// Mock of FB_AzimuthControl for the telescope state machine tests (MONETcommon#36, BROTLib plan 2026-10-21-telescope-state-machine-unification D1).
FUNCTION_BLOCK FB_AzimuthMock EXTENDS HalfBROT.FB_AzimuthControl
VAR_INPUT
	nMockMoveScans	: UINT := 60;	// scans a move takes (the telescope sees Busy meanwhile)
	bMockLatchTarget	: BOOL;	// 2026-11-11: a move ends at the target of its start (like MC_MoveAbsolute), not at the current one
	fMockFollowingError	: LREAL;	// #267: deg the encoder lags the NC set position (ActualPosition = SetPosition - this); 0 = none
	nMockStopScans	: UINT := 3;	// scans an MC_Stop takes until Done
	nMockHomeScans	: UINT := 3;	// scans a homing takes
	nMockDisableScans	: UINT := 1;	// scans MC_ExtSetPointGenDisable takes (BROTLib#101)
	bMockBrakeGate	: BOOL;			// #277: TRUE = the NC enable needs bBrakeOpen, as the real block (the rig); FALSE = the standalone mock tests
END_VAR
VAR_OUTPUT
	nStopEdges		: UINT;			// stop requests the telescope made (rising edges of StopAxis)
	nExtErrors		: UINT;			// stop or move requests that met the external setpoint generator (0x4257)
	nResetEdges		: UINT;			// resets the telescope sent to the axis (Reset())
END_VAR
VAR
	fbCore	: FB_AxisMockCore;
	pBool	: POINTER TO BOOL;
	pLreal	: POINTER TO LREAL;
	bInjected	: BOOL;
	bMockPowerLost	: BOOL;		// #232: drive power cut while bEnable stays (NC state Disabled), set with SetPowerLost
	nInjectedId	: UDINT;
	fbMockHold	: HalfBROT.FB_BrakeCloseHold;	// #277: the real hold of HalfBROT, behind the mock brake gate
	bMockEnable	: BOOL;			// the enable the mock core gets
END_VAR

// No SUPER^(): the real body (MC_* blocks, AXIS_REF) does not run. The real property setters (MoveAxis -> fbAxis.MoveTo(),
// StopAxis -> fbAxis.Stop(), HomeAxis -> _StartHoming) stay, so the telescope sees the real command interface. The model
// is driven by the levels the telescope writes and writes what the telescope reads: the base outputs and, through pointers
// (FB_Axis outputs are not writable from outside), the nested fbAxis outputs.
// #277: the real block gives the NC enable only while the brake is open (bEnable AND bAtRest AND bBrakeOpen; at rest is not
// modelled) and keeps it for the stop of a moving axis when the brake closes (HalfBROT.FB_BrakeCloseHold, the real block)
bMockEnable := bEnable;
IF bMockBrakeGate THEN
	fbMockHold(bEnable := bEnable, bBrakeEnable := bEnable AND bBrakeOpen,
		bMoving := fbCore.bInMotion OR fbCore.bTrackActive OR fbCore.bCoast OR fbCore.bStopping,	// as HalfBROT: InMotion OR Stopping
		tMaxHold := tBrakeCloseHold);
	bMockEnable := fbMockHold.bAxisEnable;
END_IF
fbCore(bEnable := bMockEnable, bPowerLost := bMockPowerLost, bHome := bHomeAxis, bMove := bMoveAxis, bStop := bStopAxis, fTarget := fPosition, fHomePosition := fCalibPosition,
	bTracking := bTracking, bLatchTarget := bMockLatchTarget, nMoveScans := nMockMoveScans, nStopScans := nMockStopScans, nHomeScans := nMockHomeScans,
	nDisableScans := nMockDisableScans);

pBool := ADR(fbAxis.Ready);			pBool^ := fbCore.bReady;
pBool := ADR(fbAxis.Calibrated);	pBool^ := fbCore.bCalibrated;
pBool := ADR(fbAxis.HomeDone);		pBool^ := fbCore.bCalibrated;
pBool := ADR(fbAxis.HomeActive);	pBool^ := fbCore.bHoming;
pBool := ADR(fbAxis.Homing);		pBool^ := fbCore.bHoming;
pBool := ADR(fbAxis.InMotion);		pBool^ := fbCore.bInMotion OR fbCore.bTrackActive OR fbCore.bCoast;
pBool := ADR(fbAxis.isTracking);	pBool^ := fbCore.bTrackActive;
pBool := ADR(fbAxis.StandStill);	pBool^ := fbCore.bStandStill AND NOT fbCore.bTrackActive AND NOT fbCore.bCoast;
pBool := ADR(fbAxis.MoveDone);		pBool^ := fbCore.bMoveDone;
pBool := ADR(fbAxis.Stopping);		pBool^ := fbCore.bStopping;
pBool := ADR(fbAxis.StopDone);		pBool^ := fbCore.bStopDone;
pBool := ADR(fbAxis.Busy);			pBool^ := fbCore.bInMotion OR fbCore.bHoming;
pLreal := ADR(fbAxis.ActualPosition);	pLreal^ := fbCore.fPosition - fMockFollowingError;
pLreal := ADR(fbAxis.SetPosition);		pLreal^ := fbCore.fPosition;	// the model position is the NC set position (#267)

bReady := fbCore.bReady AND fbCore.bStandStill;
bCalibrated := fbCore.bCalibrated;
fActualPosition := fbCore.fPosition - fMockFollowingError;
nStopEdges := fbCore.nStopEdges;
nExtErrors := fbCore.nExtErrors;
IF fbCore.bExtError THEN
	bInjected := TRUE;
	nInjectedId := 16#4257;	// Motion commands are not allowed for external setpoint generated axis
END_IF

// the real control body clears the levels like this: the move on MoveDone, the stop on StopDone, the homing request
// once the axis is calibrated and the homing procedure is over
IF fbCore.bMoveDone THEN
	bMoveAxis := FALSE;
END_IF
IF fbCore.bStopDone THEN
	bStopAxis := FALSE;
END_IF
IF fbCore.bCalibrated AND NOT fbCore.bHoming THEN
	bHomeAxis := FALSE;
END_IF
IF bReset THEN
	nResetEdges := nResetEdges + 1;
	bReset := FALSE;	// ResetDone at once
	bInjected := FALSE;
END_IF
bError := bInjected;
nErrorID := nInjectedId;

// the limit inputs the pendant reads (InDigitalInputs, AT%I*): bit 0 and 1 TRUE = limit switch free (FB_MonetPendantControl_Tests)
METHOD SetDigitalInputs
VAR_INPUT
	nInputs	: WORD;
END_VAR
InDigitalInputs := nInputs;
END_METHOD

// the axis reports an error with this id until the telescope resets it (bError/nErrorID are what the telescope reads)
METHOD InjectError
VAR_INPUT
	nId	: UDINT;
END_VAR
bInjected := TRUE;
nInjectedId := nId;
END_METHOD

// #232: the drive power is cut though the request stays (HalfBROT brake interlock): Ready and StandStill FALSE, like the NC state Disabled
METHOD SetPowerLost
VAR_INPUT
	bLost	: BOOL;
END_VAR
bMockPowerLost := bLost;
END_METHOD

END_FUNCTION_BLOCK

(* stored: Version 1.1.0.1, ProductVersion 3.1.4024.15
   POU FB_AzimuthMock: Id {f2ffd774-8a4d-4067-a41a-a990b1c8eab7}, SpecialFunc None
   Method SetDigitalInputs: Id {50c2fec9-4cfc-4444-8dec-43a084c75f72}
   Method InjectError: Id {7b5ffe42-4f43-4d92-9ec6-dd005695327d}
   Method SetPowerLost: Id {2c4a888a-544d-494f-b3c3-109fceaee724} *)
